FUNCTION_BLOCK Sensor_Generico (* Sensor analogico generico (4-20 mA ou comunicacao) - HidrycoLib *)
  (* Standard: 61499-2 *)
  (* Version 2.4, 12/11/2026, Hidryco, Hidryco, 2.4: aviso e erro do proprio dispositivo (symlinks stsAvisoDispositivo e stsErroDispositivo, INT, so com cfgComunicacao): erro = falha do sensor, aviso = alarme AlarmeAviso (Warning); codigos no diagnostico (fpParameter). 2.3: cfgSkid (valor ja escalado no skid): sensor sempre habilitado (Logica) e IHM sem escala e sem ajustes (CFG_SKID). 2.2: cfgFalhaMin/Max padrao 3800/22000 (eram 3600/21000). 2.1: saidas stsAtivoHH/stsAtivoH (alarme com tempo e sem memoria) e stsDisponivel no CNF. 2.0: tags da IO List da Nereda no IThis: CommonError (mesma origem do STS_FALHA_SENSOR), Reliability = 80 fixo e DaysToMaintenance = 0. 1.9: limites dos alarmes em unidade de engenharia (Logica.stsLimHH..LL) para o grafico da IHM. 1.8: tag STS_FALHA renomeada para STS_FALHA_SENSOR (mesmo ID F96D4140FF4E3BE0), so com a falha do sensor (fora da faixa ou falha do instrumento); a comunicacao fica em STS_FALHA_COMUNICACAO; STS_FALHA_ATIVA com qualquer falha. 1.7: E_CYCLE TickHmi (1 s): valores para a IHM no maximo 1 vez por segundo. 1.6: tag STS_FALHA_SENSOR renomeada para STS_FALHA = falha ativa (sensor em falha agora, sem memoria); nova tag STS_FALHA_COMUNICACAO (sensores por comunicacao ou com status da conexao). 1.5: sensor de nivel (cfgNivel) com os setpoints de alarme em % da altura maxima. 1.4: sinal em falha tambem pelo status da conexao Modbus (symlink stsConexao INT, 1 = online) com cfgUsaConexao, no 4-20 mA lido por remota e na comunicacao. 1.3: entrada inibeAlarmesBaixos (E_INIBE) e saidas stsCondicaoHH/H/L/LL (limite ultrapassado agora). 1.2: alarmes na lista do EAE com reconhecimento pelo reset e pisca na IHM (ISA-101), tempo padrao de alarme 5 s. 1.0: sensor generico (substitui Sensor_4a20, Sensor_Nivel_4a20 e Sensor_Comunicacao). Campo por symlink ${PATH}: 4-20 mA = stsSensorBruto (INT); comunicacao = stsFalhaSensor, stsEntrada (REAL), stsFalhaComunicacao. Alarmes HH/H/L/LL e falha no sistema de alarmes do EAE (ALARM_BIT). *)
  PACKAGE Hidryco.HidrycoLib;
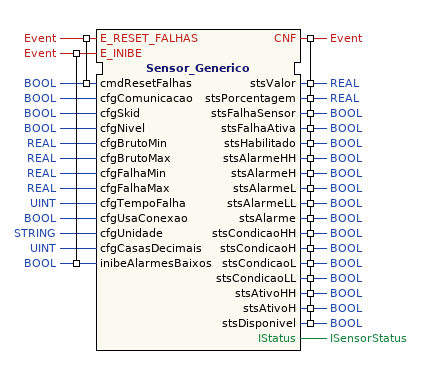
  EVENT_INPUT
    E_RESET_FALHAS WITH cmdResetFalhas; (* Reset da falha e dos alarmes pelo processo (com cmdResetFalhas = TRUE) *)
    E_INIBE WITH inibeAlarmesBaixos; (* Inibicao dos alarmes L e LL pelo processo *)
  END_EVENT
  EVENT_OUTPUT
    CNF WITH stsValor, stsPorcentagem, stsFalhaSensor, stsFalhaAtiva, stsHabilitado, stsAlarmeHH, stsAlarmeH, stsAlarmeL, stsAlarmeLL, stsAlarme, stsCondicaoHH, stsCondicaoH, stsCondicaoL, stsCondicaoLL, stsAtivoHH, stsAtivoH, stsDisponivel; (* Status (so na mudanca) *)
  END_EVENT
  VAR_INPUT
    cmdResetFalhas : BOOL; (* TRUE = reset (com o evento E_RESET_FALHAS) *)
    cfgComunicacao : BOOL := FALSE; (* FALSE = entrada 4-20 mA (stsSensorBruto), TRUE = valor por comunicacao (stsEntrada, ja em unidade de engenharia) *)
    cfgSkid : BOOL := FALSE; (* TRUE = valor vem de um skid (gradeamento, UCT, C-Press) ja escalado no proprio skid: a IHM nao mostra o ajuste de escala *)
    cfgNivel : BOOL := FALSE; (* TRUE = sensor de nivel: calcula % sobre a altura maxima *)
    cfgBrutoMin : REAL := 4000.0; (* Valor bruto em 4 mA (TM3: 4000) *)
    cfgBrutoMax : REAL := 20000.0; (* Valor bruto em 20 mA (TM3: 20000) *)
    cfgFalhaMin : REAL := 3800.0; (* Abaixo deste bruto = falha (3,8 mA) *)
    cfgFalhaMax : REAL := 22000.0; (* Acima deste bruto = falha (22,0 mA) *)
    cfgTempoFalha : UINT := 5; (* Tempo para confirmar a falha do sinal (s) *)
    cfgUsaConexao : BOOL := FALSE; (* TRUE = sinal em falha tambem quando o status da conexao Modbus (symlink stsConexao, INT: 1 = online) for diferente de 1 (4-20 mA lido por remota ou comunicacao) *)
    cfgUnidade : STRING := ''; (* Unidade de engenharia mostrada na IHM (ex.: m, bar, m3/h, mg/L) *)
    cfgCasasDecimais : UINT := 2; (* Casas decimais do valor na IHM *)
    inibeAlarmesBaixos : BOOL := FALSE; (* TRUE = alarmes L e LL inibidos (com o evento E_INIBE). Ex.: pressao de recalque com as bombas paradas *)
  END_VAR
  VAR_OUTPUT
    stsValor : REAL; (* Valor em unidade de engenharia (0 em falha ou desabilitado) *)
    stsPorcentagem : REAL; (* Nivel em % da altura maxima (so cfgNivel) *)
    stsFalhaSensor : BOOL; (* Falha do sensor memorizada (ate o reset) *)
    stsFalhaAtiva : BOOL; (* Sinal em falha agora (valor invalido) *)
    stsHabilitado : BOOL; (* Sensor habilitado *)
    stsAlarmeHH : BOOL; (* Alarme HH (memorizado ate o reset; suprimido com o sinal em falha) *)
    stsAlarmeH : BOOL; (* Alarme H (memorizado ate o reset; suprimido com o sinal em falha) *)
    stsAlarmeL : BOOL; (* Alarme L (memorizado ate o reset; suprimido com o sinal em falha) *)
    stsAlarmeLL : BOOL; (* Alarme LL (memorizado ate o reset; suprimido com o sinal em falha) *)
    stsAlarme : BOOL; (* Algum alarme ativo *)
    stsCondicaoHH : BOOL; (* Valor alem do setpoint HH agora (sem tempo e sem memoria; so com o alarme habilitado e o sinal bom) *)
    stsCondicaoH : BOOL; (* Valor alem do setpoint H agora (sem tempo e sem memoria; so com o alarme habilitado e o sinal bom) *)
    stsCondicaoL : BOOL; (* Valor alem do setpoint L agora (sem tempo e sem memoria; so com o alarme habilitado e o sinal bom) *)
    stsCondicaoLL : BOOL; (* Valor alem do setpoint LL agora (sem tempo e sem memoria; so com o alarme habilitado e o sinal bom) *)
    stsAtivoHH : BOOL; (* Alarme HH com o tempo do alarme e sem memoria (some quando o valor volta) *)
    stsAtivoH : BOOL; (* Alarme H com o tempo do alarme e sem memoria (some quando o valor volta) *)
    stsDisponivel : BOOL; (* Sensor habilitado, com leitura e sem falha *)
  END_VAR
  PLUGS
    IStatus : ISensorStatus;
  END_PLUGS
  FBS
    CampoAviso : SYMLINKMULTIVARDST_5A03F112CD5D470(NAME1 := '$${PATH}stsAvisoDispositivo'); {SET_ATTRIBUTE(Configuration.GenericFBType.InterfaceParams, Runtime.System#I:=1;VALUE${I$}:INT)}
    CampoErro : SYMLINKMULTIVARDST_5A03F112CD5D470(NAME1 := '$${PATH}stsErroDispositivo'); {SET_ATTRIBUTE(Configuration.GenericFBType.InterfaceParams, Runtime.System#I:=1;VALUE${I$}:INT)}
    AlarmeAviso : ALARM_BIT(TYPE := 1, ACKTYPE_1 := 2, ACTIVE := TRUE); {SET_ATTRIBUTE(HMI.AlarmText, Aviso do próprio sensor)} {SET_ATTRIBUTE(HMI.AlarmClass, Warning)}
    IThis : Sensor_Generico_HMI(QI := TRUE, Reliability := 80);
    plcStart1 : plcStart(Prio := 10);
    Logica : basicSensorGenerico;
    CampoBruto : SYMLINKMULTIVARDST_5A03F112CD5D470(NAME1 := '$${PATH}stsSensorBruto'); {SET_ATTRIBUTE(Configuration.GenericFBType.InterfaceParams, Runtime.System#I:=1;VALUE${I$}:INT)}
    CampoComunicacao : SYMLINKMULTIVARDST_804524063F215924(NAME1 := '$${PATH}stsFalhaSensor', NAME2 := '$${PATH}stsEntrada', NAME3 := '$${PATH}stsFalhaComunicacao'); {SET_ATTRIBUTE(Configuration.GenericFBType.InterfaceParams, Runtime.System#I:=3;VALUE${I$}:BOOL,REAL,BOOL)}
    CampoConexao : SYMLINKMULTIVARDST_5A03F112CD5D470(NAME1 := '$${PATH}stsConexao'); {SET_ATTRIBUTE(Configuration.GenericFBType.InterfaceParams, Runtime.System#I:=1;VALUE${I$}:INT)}
    DelayFalha : E_DELAY;
    DelayHH : E_DELAY;
    DelayH : E_DELAY;
    DelayL : E_DELAY;
    DelayLL : E_DELAY;
    AlarmeHH : ALARM_BIT(TYPE := 1, ACKTYPE_1 := 2, ACTIVE := TRUE); {SET_ATTRIBUTE(HMI.AlarmText, Medição muito alta (HH))}
    AlarmeH : ALARM_BIT(TYPE := 1, ACKTYPE_1 := 2, ACTIVE := TRUE); {SET_ATTRIBUTE(HMI.AlarmText, Medição alta (H))} {SET_ATTRIBUTE(HMI.AlarmClass, Warning)}
    AlarmeL : ALARM_BIT(TYPE := 1, ACKTYPE_1 := 2, ACTIVE := TRUE); {SET_ATTRIBUTE(HMI.AlarmText, Medição baixa (L))} {SET_ATTRIBUTE(HMI.AlarmClass, Warning)}
    AlarmeLL : ALARM_BIT(TYPE := 1, ACKTYPE_1 := 2, ACTIVE := TRUE); {SET_ATTRIBUTE(HMI.AlarmText, Medição muito baixa (LL))}
    AlarmeFalha : ALARM_BIT(TYPE := 1, ACKTYPE_1 := 2, ACTIVE := TRUE); {SET_ATTRIBUTE(HMI.AlarmText, Falha do sensor ou do sinal)}
    TickHmi : E_CYCLE(DT := T#1s);
  END_FBS
  EVENT_CONNECTIONS
    plcStart1.FIRST_INIT TO IThis.B11E9EDFB330BB0A;
    plcStart1.REDO_INIT TO IThis.B11E9EDFB330BB0A;
    IThis.8DA9E22D0BD63DE1 TO Logica.A313A1584C9E1BE5;
    Logica.AFC15B7A52538DC1 TO CampoBruto.INIT;
    Logica.AFC15B7A52538DC1 TO CampoComunicacao.INIT;
    Logica.AFC15B7A52538DC1 TO AlarmeHH.INIT;
    AlarmeHH.INITO TO AlarmeHH.REQ_INITDATA;
    AlarmeHH.CNF_INITDATA TO AlarmeHH.ACTIVATE;
    AlarmeHH.INITO TO AlarmeH.INIT;
    AlarmeH.INITO TO AlarmeH.REQ_INITDATA;
    AlarmeH.CNF_INITDATA TO AlarmeH.ACTIVATE;
    AlarmeH.INITO TO AlarmeL.INIT;
    AlarmeL.INITO TO AlarmeL.REQ_INITDATA;
    AlarmeL.CNF_INITDATA TO AlarmeL.ACTIVATE;
    AlarmeL.INITO TO AlarmeLL.INIT;
    AlarmeLL.INITO TO AlarmeLL.REQ_INITDATA;
    AlarmeLL.CNF_INITDATA TO AlarmeLL.ACTIVATE;
    AlarmeLL.INITO TO AlarmeFalha.INIT;
    AlarmeFalha.INITO TO AlarmeFalha.REQ_INITDATA;
    AlarmeFalha.CNF_INITDATA TO AlarmeFalha.ACTIVATE;
    AlarmeFalha.INITO TO plcStart1.ACK_FIRST;
    AlarmeFalha.INITO TO IThis.F46E32F8CF51BE9D;
    CampoBruto.CNF TO Logica.BB3A40EF748E4AD2;
    CampoComunicacao.CNF TO Logica.85BF8544E9C17F76;
    IThis.BC1F18854FDB14ED TO Logica.60FC42EE781F51CC;
    IThis.4275246E291683C0 TO Logica.2394F0A61CB1494A;
    E_RESET_FALHAS TO Logica.20033B1C8F10344F;
    E_INIBE TO Logica.F6476A371C298363;
    IStatus.9E548C371B42FEDC TO Logica.C81E4D5CD6D5669B;
    Logica.8A583D6DDA99E174 TO DelayFalha.STOP;
    Logica.88B29E7FCEDFD04A TO DelayFalha.START;
    DelayFalha.EO TO Logica.79D90CC239980ABE;
    Logica.AC54F201197F1308 TO DelayHH.STOP;
    Logica.AD777C25E731B753 TO DelayHH.START;
    DelayHH.EO TO Logica.0507438F316FE05A;
    Logica.600AE8762D264606 TO DelayH.STOP;
    Logica.286E3580B6A4E911 TO DelayH.START;
    DelayH.EO TO Logica.60C0262360B78E5E;
    Logica.64E82BD205C26648 TO DelayL.STOP;
    Logica.A5C367FB8CC6123F TO DelayL.START;
    DelayL.EO TO Logica.2ED9A6722EA41B53;
    Logica.F8318F17CCD7636C TO DelayLL.STOP;
    Logica.48A9F0D2C448300B TO DelayLL.START;
    DelayLL.EO TO Logica.1B3FD32E01035504;
    Logica.AD639990F05475A6 TO CNF;
    Logica.FC4E06ABE3EBBDDF TO IStatus.C09F18F0C837B93D;
    Logica.ABC9F934A736FB9D TO IStatus.AB5911D326737849;
    Logica.4113A4030DCFA861 TO IThis.0DB49FB1D65E52DB;
    Logica.DA3C0D9212A1D794 TO AlarmeHH.REQ;
    Logica.DA3C0D9212A1D794 TO AlarmeH.REQ;
    Logica.DA3C0D9212A1D794 TO AlarmeL.REQ;
    Logica.DA3C0D9212A1D794 TO AlarmeLL.REQ;
    Logica.DA3C0D9212A1D794 TO AlarmeFalha.REQ;
    AlarmeHH.IND_1 TO IThis.0DB49FB1D65E52DB;
    AlarmeH.IND_1 TO IThis.0DB49FB1D65E52DB;
    AlarmeL.IND_1 TO IThis.0DB49FB1D65E52DB;
    AlarmeLL.IND_1 TO IThis.0DB49FB1D65E52DB;
    AlarmeFalha.IND_1 TO IThis.0DB49FB1D65E52DB;
    IThis.4275246E291683C0 TO AlarmeHH.ACK_C1;
    IThis.4275246E291683C0 TO AlarmeH.ACK_C1;
    IThis.4275246E291683C0 TO AlarmeL.ACK_C1;
    IThis.4275246E291683C0 TO AlarmeLL.ACK_C1;
    IThis.4275246E291683C0 TO AlarmeFalha.ACK_C1;
    Logica.AFC15B7A52538DC1 TO CampoConexao.INIT;
    CampoConexao.CNF TO Logica.BA1EF67945330BA4;
    Logica.AFC15B7A52538DC1 TO TickHmi.START;
    TickHmi.EO TO Logica.01B9A26CA80ECAC9;
    Logica.AFC15B7A52538DC1 TO CampoAviso.INIT;
    Logica.AFC15B7A52538DC1 TO CampoErro.INIT;
    CampoAviso.CNF TO Logica.13DE6C7C018FFF3E;
    CampoErro.CNF TO Logica.13DE6C7C018FFF3E;
    AlarmeFalha.INITO TO AlarmeAviso.INIT;
    AlarmeAviso.INITO TO AlarmeAviso.REQ_INITDATA;
    AlarmeAviso.CNF_INITDATA TO AlarmeAviso.ACTIVATE;
    Logica.DA3C0D9212A1D794 TO AlarmeAviso.REQ;
    AlarmeAviso.IND_1 TO IThis.0DB49FB1D65E52DB;
    IThis.4275246E291683C0 TO AlarmeAviso.ACK_C1;
  END_CONNECTIONS
  DATA_CONNECTIONS
    cfgComunicacao TO Logica.BDC9951972159B49;
    cfgNivel TO Logica.A121066C0B4E396A;
    cfgBrutoMin TO Logica.08668FFBD0D4C224;
    cfgBrutoMax TO Logica.5C5752CDF95E2D99;
    cfgFalhaMin TO Logica.D75E79B6B7019547;
    cfgFalhaMax TO Logica.E942EB878618E7C8;
    cfgTempoFalha TO Logica.2D81E0FCE9B8E921;
    cmdResetFalhas TO Logica.A71A8E7BCD5DEA8F;
    IStatus.E54954E6518AFFE0 TO Logica.A114BF4DF6C8FACD;
    inibeAlarmesBaixos TO Logica.CB16E6E7444E9F47;
    Logica.0D31DC1406BFACF0 TO CampoBruto.QI;
    Logica.9DEE58A20A0B0AFD TO CampoComunicacao.QI;
    CampoBruto.VALUE1 TO Logica.AF52988DC4E16721;
    CampoComunicacao.VALUE1 TO Logica.DC02530AB13A0CE9;
    CampoComunicacao.VALUE2 TO Logica.127AA48C83FCE0F9;
    CampoComunicacao.VALUE3 TO Logica.AC6220939047FF1C;
    Logica.1F6F64330B9EFE72 TO DelayFalha.DT;
    Logica.F3031E01158FE3E1 TO DelayHH.DT;
    Logica.585F9BC133BAE667 TO DelayH.DT;
    Logica.AFF40B3AA17C5F37 TO DelayL.DT;
    Logica.D17EC1927CB7668B TO DelayLL.DT;
    IThis.74F7308C27744D49 TO Logica.BCFBEA21C064840B;
    IThis.0BD1CDAA1517CE9D TO Logica.1EF616CE5E6D0F0D;
    IThis.80A8E9E8A637C9EC TO Logica.A67F7A68A4947959;
    IThis.9F16D125566454DD TO Logica.40810CB570D37DC2;
    IThis.93AF73B64660FBA6 TO Logica.093F317F91681B94;
    IThis.A8AE53BDCD5D904B TO Logica.2368E646122F6C1E;
    IThis.D202A579D84D6111 TO Logica.61BA9A4108167FE1;
    IThis.D0AF2971D81905DB TO Logica.E7EC039942CE430E;
    IThis.7654A9844654582E TO Logica.44FFB666822352BF;
    IThis.9F33F2002C72AA38 TO Logica.1B30B39C75AABA90;
    IThis.20FFBF6BD7638BE5 TO Logica.3B12D5C113628B3D;
    IThis.27BF8C3F14711ABA TO Logica.0C17F55C15BCD39D;
    IThis.81B00D22F26005A0 TO Logica.275E0286C790B3B5;
    IThis.CA2F98887484603A TO Logica.91055F2FEA3A7CFE;
    IThis.CC9F410D4B3B3695 TO Logica.5837C50851352086;
    IThis.5C9A19D23397D700 TO Logica.43D87B8E2D957E3F;
    IThis.23C877B7D5B67937 TO Logica.12DA5CE2186CD3E9;
    Logica.7CD1C7E9D29D5BA8 TO AlarmeHH.INP;
    Logica.2175D6B4C45D9235 TO AlarmeH.INP;
    Logica.D792B1098650EBBE TO AlarmeL.INP;
    Logica.123CA78819C21E67 TO AlarmeLL.INP;
    Logica.9751C9BCFBC02314 TO AlarmeFalha.INP;
    Logica.3203282664F84EE7 TO stsValor;
    Logica.E36A36073A4D8255 TO stsPorcentagem;
    Logica.D2CE0143DEEF5F5B TO stsFalhaSensor;
    Logica.90D219EA9609F475 TO stsFalhaAtiva;
    Logica.BC2F73C5CA9874F4 TO stsHabilitado;
    Logica.846DCED7A53DAF52 TO stsAlarmeHH;
    Logica.11F28407C39B0DB4 TO stsAlarmeH;
    Logica.41F92ED47B97DD7B TO stsAlarmeL;
    Logica.F2CABDC5ADA79A97 TO stsAlarmeLL;
    Logica.478DE584A3EC80F6 TO stsAlarme;
    Logica.5C7B1A72AEA1734C TO stsCondicaoHH;
    Logica.B271C2D0A9370A7F TO stsCondicaoH;
    Logica.80C046EE3841337A TO stsCondicaoL;
    Logica.46248A230C3897E2 TO stsCondicaoLL;
    Logica.3203282664F84EE7 TO IThis.8897CDA500AC3B43;
    Logica.E36A36073A4D8255 TO IThis.03F005FFEA8B1EB7;
    Logica.821A07A8E8DE848B TO IThis.8C3B32492EDE30F6;
    Logica.D2CE0143DEEF5F5B TO IThis.F96D4140FF4E3BE0;
    Logica.D2CE0143DEEF5F5B TO IThis.339076CC42EE7FBD;
    Logica.90D219EA9609F475 TO IThis.50692E037DBEB5AF;
    Logica.81E22B6ADE19C4D7 TO IThis.3066A0DA727B2781;
    Logica.BC2F73C5CA9874F4 TO IThis.8CC7DAAF94A2F272;
    Logica.846DCED7A53DAF52 TO IThis.F359F702D2084BBB;
    Logica.11F28407C39B0DB4 TO IThis.A44C5B0C739C913A;
    Logica.41F92ED47B97DD7B TO IThis.02D192408DD0BAD7;
    Logica.F2CABDC5ADA79A97 TO IThis.383A34199F936BCE;
    Logica.478DE584A3EC80F6 TO IThis.D2378FEEF5A3D1D1;
    Logica.8550C71DBEEC8F3F TO IThis.D7B779974D991A8E;
    cfgComunicacao TO IThis.CBCE958A8B6D12A1;
    cfgNivel TO IThis.8BC973C9232A9202;
    cfgUnidade TO IThis.1A77C34E03AFA0CE;
    cfgCasasDecimais TO IThis.4834B2F21AEC2CC6;
    AlarmeHH.STATE_1 TO IThis.A91C3C65B4F67DE5;
    AlarmeH.STATE_1 TO IThis.B10CA9D36B32EBC9;
    AlarmeL.STATE_1 TO IThis.02DAB08BEDD4D70F;
    AlarmeLL.STATE_1 TO IThis.C4A67D01408D3D56;
    AlarmeFalha.STATE_1 TO IThis.D31A79F7D2BBEF19;
    Logica.3203282664F84EE7 TO IStatus.BC22E5B309EC3525;
    Logica.90D219EA9609F475 TO IStatus.C4FED0E2B2BCAFA9;
    Logica.846DCED7A53DAF52 TO IStatus.7C32AA46813E72EF;
    Logica.11F28407C39B0DB4 TO IStatus.1A87F8257AB469E4;
    Logica.41F92ED47B97DD7B TO IStatus.F1DB93298B22A3D1;
    Logica.F2CABDC5ADA79A97 TO IStatus.D6ADC459B9EEBD4A;
    cfgUsaConexao TO Logica.5A40623945DBD51C;
    Logica.DD2B06522C2E1D6D TO CampoConexao.QI;
    CampoConexao.VALUE1 TO Logica.A01E732EBCA193E3;
    Logica.72AFED77258A9210 TO IThis.4D0002C974B24A69;
    Logica.082D88F711CCD739 TO IThis.2007E90E21C8B4CF;
    Logica.D91E42414EEE194E TO IThis.7B165BE1315191C3;
    Logica.6D7F45595C9C84C3 TO IThis.FFEA0503A1019B14;
    Logica.1C96D9FB2C39CC10 TO stsAtivoHH;
    Logica.48B250C8BC490C7B TO stsAtivoH;
    Logica.0DF0DDE240BFC12B TO stsDisponivel;
    cfgSkid TO IThis.BB5D27FFFC44E39C;
    cfgSkid TO Logica.C03D96BA9EA046E5;
    Logica.9DEE58A20A0B0AFD TO CampoAviso.QI;
    Logica.9DEE58A20A0B0AFD TO CampoErro.QI;
    CampoAviso.VALUE1 TO Logica.DB454D1BA11A0DE9;
    CampoErro.VALUE1 TO Logica.222F1372FEE9B05F;
    Logica.789D37109634E4C8 TO AlarmeAviso.INP;
    AlarmeAviso.STATE_1 TO IThis.F428A55205D49D87;
    Logica.7DE82A7B3D5EBDF3 TO IThis.8291008A357A190E;
    Logica.CC00142E36E22C6A TO IThis.F79BEE55D150EAB5;
  END_CONNECTIONS
END_FUNCTION_BLOCK
